// TIA Portal V21 export
// export: Created 2026-11-10T07:35:09.7637249Z, ExportSetting WithDefaults, DisplayName Totally Integrated Automation Portal, DisplayVersion V21 Update 3, DisplayName STEP 7 Professional, DisplayVersion V21 Update 3, DisplayName STEP 7 Safety, DisplayVersion V21, DisplayName Tech WebApplication, DisplayVersion V21, DisplayName WinCC Basic/Comfort/Advanced, DisplayVersion V21 Update 3, DisplayName WinCC Unified, DisplayVersion V21 Update 3
FUNCTION_BLOCK "FB_Lad_ex094"   // FB188, LAD
{ S7_Optimized_Access := 'TRUE' }
VERSION : 0.1
// stored: AutoNumber true, IsIECCheckEnabled false, IsRetainMemResEnabled false, MemoryReserve 100, SetENOAutomatically false, UDAEnableTagReadback false
   VAR_INPUT
      v_pe_i_dev_new : Bool;
      v_cmd : Int;
      v_cmd_modifier : Int;
      v_count : Byte;
   END_VAR
   VAR_OUTPUT
      v_error : Bool;
      v_status : Word;
   END_VAR
   VAR_IN_OUT
      v_activate : Bool;
      v_valid : Bool;
      v_measurement_list : Variant;
      v_data_errorrsp : Variant;
   END_VAR
BEGIN

REGION Network 1: PE_Measurement_List_RSP - Generate list of supported measured values as answer
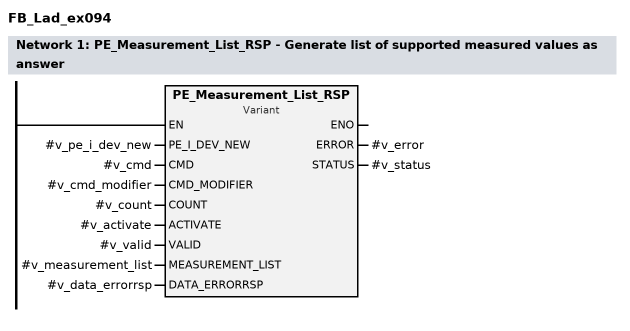
   RUNG wire#powerrail
      { S7_Templates := "[data_errorrsp_type := Variant, measurement_list_type := Variant]" } PE_Measurement_List_RSP(PE_I_DEV_NEW := #v_pe_i_dev_new, CMD := #v_cmd, CMD_MODIFIER := #v_cmd_modifier, Count := #v_count, Activate := #v_activate, VALID := #v_valid, ERROR => #v_error, STATUS => #v_status, Measurement_List := #v_measurement_list, DATA_ERRORRSP := #v_data_errorrsp)
   END_RUNG
   // the same network as SCL:
   PE_Measurement_List_RSP(PE_I_DEV_NEW := #v_pe_i_dev_new,
                           CMD := #v_cmd,
                           CMD_MODIFIER := #v_cmd_modifier,
                           Count := #v_count,
                           Activate := #v_activate,
                           VALID := #v_valid,
                           Measurement_List := #v_measurement_list,
                           DATA_ERRORRSP := #v_data_errorrsp,
                           ERROR => #v_error,
                           STATUS => #v_status);
END_REGION
END_FUNCTION_BLOCK
